Fanuc KAREL source: kt00074.KL

-- PROVISIONAL review KL for V1013-1; original PC SHA256 02506bf35f5e20fae9f9d1e9de0ec900d835ee32518129e0bbbacab8daf3f4c7
-- Incomplete behavior may be omitted. Consult companion uncertainty JSON. Do not deploy.
PROGRAM KT00074
%NOLOCKGROUP
VAR
  R1 : REAL
  I2 : INTEGER
  OUT : REAL
BEGIN
  -- UNRESOLVED_PC offsets 5-16; opcodes 2E,23
  -- UNRESOLVED_PC offsets 21-32; opcodes 2E,23
  -- UNRESOLVED_PC offsets 37-57; opcodes 21,21,64,6B,23
  -- UNRESOLVED_PC offsets 62-66; opcodes 7F
END KT00074
